// TIA Portal V21 export
// export: Created 2026-11-10T07:35:19.7013902Z, ExportSetting WithDefaults, DisplayName Totally Integrated Automation Portal, DisplayVersion V21 Update 3, DisplayName STEP 7 Professional, DisplayVersion V21 Update 3, DisplayName STEP 7 Safety, DisplayVersion V21, DisplayName Tech WebApplication, DisplayVersion V21, DisplayName WinCC Basic/Comfort/Advanced, DisplayVersion V21 Update 3, DisplayName WinCC Unified, DisplayVersion V21 Update 3
FUNCTION_BLOCK "FB_Lad_ex140"   // FB106, LAD
{ S7_Optimized_Access := 'TRUE' }
VERSION : 0.1
// stored: AutoNumber true, IsIECCheckEnabled false, IsRetainMemResEnabled false, MemoryReserve 100, SetENOAutomatically false, UDAEnableTagReadback false
   VAR_INPUT
      v_req : Bool;
      v_mode : UInt;
      v_name : Array[0..99] of Byte;
   END_VAR
   VAR_OUTPUT
      v_done : Bool;
      v_busy : Bool;
      v_error : Bool;
      v_status : Word;
   END_VAR
   VAR_IN_OUT
      v_id : DWord;
      v_data : Array[0..99] of Byte;
   END_VAR
   VAR
      inst { S7_SetPoint := 'True'} : DataLogOpen;
   END_VAR
BEGIN

REGION Network 1: DataLogOpen - Open data log
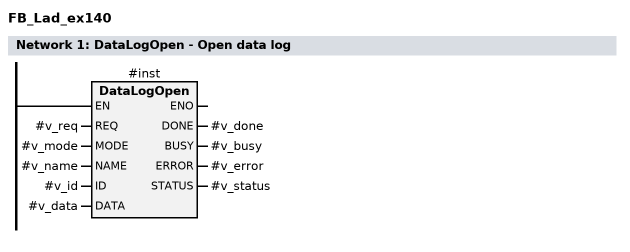
   RUNG wire#powerrail
      { S7_Templates := "card := 1" } #inst.DataLogOpen(REQ := #v_req, MODE := #v_mode, "NAME" := #v_name, ID := #v_id, Data := #v_data, DONE => #v_done, BUSY => #v_busy, ERROR => #v_error, STATUS => #v_status)
   END_RUNG
   // the same network as SCL:
   #inst(REQ := #v_req,   // DataLogOpen
         MODE := #v_mode,
         "NAME" := #v_name,
         ID := #v_id,
         Data := #v_data,
         DONE => #v_done,
         BUSY => #v_busy,
         ERROR => #v_error,
         STATUS => #v_status);
END_REGION
END_FUNCTION_BLOCK
